(* CODESYS project winhmi.library
   DefaultNamespace: KOSTAL.AF2024.HMI.WinHMI
   DocFormat: reStructuredText
   Description: Interface to WinHMI application
   Author: Martin Hundt
   Title: KOSTAL.AF2024.HMI.WinHMI
   Version: 2.0.0.0
   Company: KOSTAL GmbH & Co.KG
   Placeholder: KOSTAL.AF2024.HMI.WinHMI

Project tree, tasks and I/O mapping:
  libraries: KOSTAL.AF2024.Core.functionResponse, 1.0.0.0 (KOSTAL GmbH & Co.KG); KOSTAL.AF2024.Core.GetSystemTime, 1.0.1.0 (KOSTAL GmbH & Co.KG); KOSTAL.AF2024.Core.ID, 1.0.0.0 (KOSTAL GmbH & Co.KG); KOSTAL.AF2024.Core.JsonTools, 1.0.0.0 (KOSTAL GmbH & Co.KG); KOSTAL.AF2024.Core.ListOf, 1.0.0.0 (KOSTAL GmbH & Co.KG); KOSTAL.AF2024.Core.MainControl, 1.0.0.0 (KOSTAL GmbH & Co.KG); KOSTAL.AF2024.Core.Process, 1.0.999.1 (KOSTAL GmbH & Co.KG); KOSTAL.AF2024.Core.Settings, 1.0.0.0 (KOSTAL GmbH & Co.KG); KOSTAL.AF2024.Core.Station, 1.0.0.0 (KOSTAL GmbH & Co.KG); KOSTAL.AF2024.Core.StringTools, 1.0.0.0 (KOSTAL GmbH & Co.KG); KOSTAL.AF2024.Core.System, 1.0.0.0 (KOSTAL GmbH & Co.KG); KOSTAL.AF2024.Core.Text, 1.0.0.0 (KOSTAL GmbH & Co.KG); KOSTAL.AF2024.HMI.Controls, 1.0.1.0 (KOSTAL GmbH & Co.KG); KOSTAL.AF2024.HMI.I_Hmi, 1.0.0.0 (KOSTAL GmbH & Co.KG); KOSTAL.AF2024.Misc.Counter, 1.0.1.0 (KOSTAL GmbH & Co.KG); Tc2_Standard, 3.4.5.0 (Beckhoff Automation GmbH); Tc2_Utilities, 3.8.2.0 (Beckhoff Automation GmbH); Tc3_JsonXml, 3.4.4.0 (Beckhoff Automation GmbH)
  Aliases/
    data type T_ARTICLESJSON
    data type T_BUTTON_LISTING
    data type T_ExpertPageUserIndex
    data type T_MEDIA_PATH
    data type T_PARAMETERJSON
    data type T_PARAMETERVALUE
  Article/
    data type _ST_Article_FromDevice
    data type _ST_Article_ToDevice
    function block FB_ArticleList [ST]: ActualArticle, AddArticle, Clear, FB_init, FBmain, SelectedArticleName, Set
    interface I_Article: ActualArticle, SelectedArticleName
  Counter/
    data type _ST_Counter_FromDevice
    data type _ST_Counter_ToDevice
    function block FB_Counter [ST]: _HMI_define, ResetEnable
  Listing/
    data type _ST_Listing_FromDevice
    data type _ST_Listing_ToDevice
    function block FB_Page_Listing [ST]: _buttonHandler, _buttonHandler_listing, _listingHandler, _setButton, FB_init, FBmain
  MainControl/
    DUT/
      ListOfIcondition/
        interface I_ListOfCondition: NumberOfMember
        interface I_ListOfCondition_Owner
      data type _E_MainControlMode
      data type _E_MainControlState
    data type _ST_MainControl_FromDevice
    data type _ST_MainControl_toDevice
    function block FB_MainControl [ST]: _buttonHandler, _mainControlHandler, _modeToEnum, _plcStateToEnum, clear, FBmain, ManualDeviceControl
    interface I_MainControl: clear
  Media/
    data type _ST_Media_ToDevice
    function block FB_Media [ST]: Clear, FBmain, SetMedia, ShowMedia, StandardPath
    interface I_Media: Clear, SetMedia, ShowMedia, StandardPath
  Parameters/
    function block _FB_jsonHandler [ST]: Clear, GetJsonString, getValue, ID, NumberOfValues, setValue, Timestamp, _Step_ClearContent, _Step_CreateContent, _Step_ParseContent
    data type _ST_Parameters_FromDevice
    data type _ST_Parameters_ToDevice
    data type E_DataMode
    function block FB_Parameters_Base [ST]: _getParameterValue, _setParameterValue, FullQualifiedFile, ReloadDataFile, _Idle, _readFile, _setParaValue, _HMIdefine, _parameterControl, _resetCondition, FBmain, link_I_getTime
  Project Information/
    function F_GetCompany [ST]
    function F_GetTitle [ST]
    function F_GetVersion [ST]
  Station/
    data type _ST_StationPage_FromDevice
    data type _ST_StationPage_ToDevice
    function block FB_Page_Station [ST]: _buttonHandler, _setButton, _stationHandler, FB_init, FBmain
  Version/
    global variables Global_Version
  XYZ/
    data type _ST_XYZ_FromDevice
    data type _ST_XYZ_ToDevice
    function block FB_page_XYZ [ST]: _buttonHandler, _fillTextLines, _pageHandler, _setButton, FB_init, FBmain
  global variables GVL_CONSTANT
*)

// Aliases/T_ARTICLESJSON
TYPE T_ARTICLESJSON : STRING(6000)
; END_TYPE

// Aliases/T_BUTTON_LISTING
TYPE T_BUTTON_LISTING : WSTRING(3); END_TYPE

// Aliases/T_ExpertPageUserIndex
(*
Description
===========
| Limited data type for the index of an expert page user
*)
TYPE T_ExpertPageUserIndex : INT(0..GVL_CONSTANT.MAX_EXPERT_STATIONS); END_TYPE

// Aliases/T_MEDIA_PATH
TYPE T_MEDIA_PATH : STRING(80)
; END_TYPE

// Aliases/T_PARAMETERJSON
TYPE T_PARAMETERJSON : STRING(6000)
; END_TYPE

// Aliases/T_PARAMETERVALUE
TYPE T_PARAMETERVALUE : STRING(40)
; END_TYPE

// Article/_ST_Article_FromDevice
(*
Description
===========
| Data type to receive article data from WinHMI display
*)
{attribute 'pack_mode' := '1'}
TYPE _ST_Article_FromDevice :
	STRUCT
		SelectedArticleName 	: T_ARTICLENAME;
	END_STRUCT
END_TYPE

// Article/_ST_Article_ToDevice
(*
Description
===========
| Data type to provide article data to WinHMI display
*)
{attribute 'pack_mode' := '1'}
TYPE _ST_Article_ToDevice :
	STRUCT
		ArticleList		: T_ARTICLESJSON;
		ActualArticle 	: T_ARTICLENAME;		(*Shows the actual used Article name	 *)
	END_STRUCT
END_TYPE

// Counter/_ST_Counter_FromDevice
(*
Description
===========
| Data type to provide counter data to WinHMI display
*)
{attribute 'pack_mode' := '1'}
TYPE _ST_Counter_FromDevice :
	STRUCT
		Reset	: BOOL;
	END_STRUCT
END_TYPE

// Counter/_ST_Counter_ToDevice
(*
Description
===========
| Data type to provide counter data to WinHMI display
*)
{attribute 'pack_mode' := '1'}
TYPE _ST_Counter_ToDevice :
	STRUCT
		Passparts		: UDINT;
		Failparts		: UDINT;
		CounterReady 	: BOOL;
		ResetEnable		: BOOL;
	END_STRUCT
END_TYPE

// Listing/_ST_Listing_FromDevice
(*
Description
===========
| Data type to receive listing page data from WinHMI display
*)
{attribute 'pack_mode' := '1'}
TYPE _ST_Listing_FromDevice :
	STRUCT
		IsActive 		: BOOL;		(* 	BOOL	-	Response the state of the Listing Form	 *)
		Button_Left	 	: ARRAY [1..GVL_CONSTANT.LISTING_MAX_LINE] OF BOOL;		(* 	ARRAY[1..10] OF BOOL	-	Status of Button - TRUE = pressed	 *)
		Button_Right	: ARRAY [1..GVL_CONSTANT.LISTING_MAX_LINE] OF BOOL;		(* 	ARRAY[1..10] OF BOOL	-	Status of Button - TRUE = pressed	 *)
	END_STRUCT
END_TYPE

// Listing/_ST_Listing_ToDevice
(*
Description
===========
| Data type to provide listing page data to WinHMI display
*)
{attribute 'pack_mode' := '1'}
TYPE _ST_Listing_ToDevice :
	STRUCT
		
		Activate 		: BOOL;		(* 	BOOL	-	Activate the Listing Form	 *)
		
		Buttons_Left_Active : WORD;		(* 	If bit is TRUE than the correspond Button is visible	 *)
		Buttons_Right_Active : WORD;		(* 	If bit is TRUE than the correspond Button is visible	 *)
		
		Buttons_Left_Text	: ARRAY [1..GVL_CONSTANT.LISTING_MAX_LINE] OF T_BUTTON_LISTING;
		Buttons_Right_Text	: ARRAY [1..GVL_CONSTANT.LISTING_MAX_LINE] OF T_BUTTON_LISTING;
		
		Text 				: ARRAY [1..GVL_CONSTANT.LISTING_MAX_LINE] OF KOSTAL_AF2024_HMI_I_Hmi.T_PAGE_TEXT;	(* Contains the Texts for Line 1..10	 *)
		Status 				: ARRAY [1..GVL_CONSTANT.LISTING_MAX_LINE] OF KOSTAL_AF2024_HMI_I_Hmi.E_STATE;		(* 	Contains the States for Line 1..10	 *)
	END_STRUCT
END_TYPE

// MainControl/DUT/_E_MainControlMode
{attribute 'qualified_only'}
{attribute 'strict'}
TYPE _E_MainControlMode :
(
	undefined := 0,	
	manual,			
	automatic
)USINT;
END_TYPE

// MainControl/DUT/_E_MainControlState
{attribute 'qualified_only'}
{attribute 'strict'}
TYPE _E_MainControlState :
(
	off := 0,	//Power off
	on,			//Power on
	calibrate,	//Power off
	ready,		//Ready to start
	busy,		//running
	finish		//Run empty
)USINT;
END_TYPE

// MainControl/_ST_MainControl_FromDevice
(*
Description
===========
| Data type to receive Main Control data from WinHMI display
*)
{attribute 'pack_mode' := '1'}
TYPE _ST_MainControl_FromDevice :
	STRUCT
		Language 			: T_LANGUAGENAME;		(* 	STRING(40)	- Selected Languagename	 *)
				
		Button_Auto 		: BOOL;		(* 	BOOL	- Status of Button - TRUE = pressed	 *)
		Button_Manual : BOOL;		(* 	BOOL	- Status of Button - TRUE = pressed	 *)
		Button_Door 		: BOOL;		(* 	BOOL	- Status of Button - TRUE = pressed	 *)

		Button_OnOff 		: BOOL;		(* BOOL *)
		Button_StartStop : BOOL;		(* BOOL *)
		Button_workEmpty : BOOL;		(* BOOL *)
		
		UserLevel	: BYTE; 	//operator = 0, service = 1, quality = 2

	END_STRUCT
END_TYPE

// MainControl/_ST_MainControl_toDevice
(*
Description
===========
| Data type to provide Main Control data to WinHMI display
*)
{attribute 'pack_mode' := '1'}
TYPE _ST_MainControl_toDevice :
	STRUCT
		Status_Auto 	: BOOL;		(* 	BOOL	-	If TRUE > Text "Auto" has a yellow background	 *)
		Status_Manual : BOOL;		(* 	BOOL	-	If TRUE > Text "Manual" has a yellow background	 *)
	
		Status_Door_Close : BOOL;		(* 	BOOL	-	If TRUE > Text "Door" has a blue background	 *)
		Status_Door_Open 	: BOOL;		(* 	BOOL	-	If TRUE > Text "Door" has a red background	 *)
		Status_Door_Safe 	: BOOL;		(* 	BOOL	-	If TRUE > Text "Door" has a green background	 *)

		Manual_Enable 	: BOOL;		(* 	BOOL	-	If TRUE > Button in bottom of Text "Manual" is visible	 *)
		Parameters_Enable 		: BOOL;		(* 	BOOL	-	If TRUE > Button in bottom of Text "Data" is visible	 *)
		Auto_Enable 		: BOOL;		(* 	BOOL	-	If TRUE > Button in bottom of Text "Auto" is visible	 *)
		Door_Enable 		: BOOL;		(* 	BOOL	-	If TRUE > Button in bottom of Text "Door" is visible	 *)
		Article_Enable 	: BOOL;		(* 	BOOL	-	If TRUE > Button in bottom of Text "Article" is visible	 *)

		(*  Buttons *)
		OnOff_Enable	: BOOL;
		RunStop_Enable	: BOOL;
		RunEmpty_Enable 	: BOOL;
		
		Status_On 		: BOOL;		(* BOOL *)
		Status_Run 		: BOOL;		(* BOOL *)
		Status_RunEmpty 	: BOOL;		(* BOOL *)
		ManualDeviceControl_Enable	: BOOL;
		
		//main Control
		State		: USINT;
		Mode		: USINT;
				
	END_STRUCT
END_TYPE

// Media/_ST_Media_ToDevice
(*
Description
===========
| Data type to provide article data to WinHMI display
*)
{attribute 'pack_mode' := '1'}
TYPE _ST_Media_ToDevice :
	STRUCT
		MediaAddress		: T_MEDIA_PATH;
	END_STRUCT
END_TYPE

// Parameters/_ST_Parameters_FromDevice
(*
Description
===========
| Data type to receive parameter data from WinHMI display
*)
{attribute 'pack_mode' := '1'}
TYPE _ST_Parameters_FromDevice :
	STRUCT
		SelectedParameter 			: BYTE;		(* 	BYTE	- Selected Dataset 	 *)
		NewValue 				: T_PARAMETERVALUE;		(* 	STRING(40)	-	New Data value	 *)
		NewValueTransmit 	: BOOL;		(* 	BOOL	-	New value is valid	 *)

	END_STRUCT
END_TYPE

// Parameters/_ST_Parameters_ToDevice
(*
Description
===========
| Data type to provide XYZ page parameter data to WinHMI display
*)
{attribute 'pack_mode' := '1'}
TYPE _ST_Parameters_ToDevice :
	STRUCT
		ParameterValuesJson		: T_PARAMETERJSON;
		NewValueAccept			: BOOL;
	END_STRUCT
END_TYPE

// Parameters/E_DataMode
{attribute 'qualified_only'}
{attribute 'strict'}
TYPE E_DataMode :
(
	Idle := 0,
	ReadFile,
	WriteParameter
);
END_TYPE

// Station/_ST_StationPage_FromDevice
(*
Description
===========
| Data type to receive 3D page from WinHMI display
*)
{attribute 'pack_mode' := '1'}
TYPE _ST_StationPage_FromDevice :
	STRUCT
		Button_F1 : BOOL;		(* 	BOOL	- Status of Button - TRUE = pressed	 *)
		Button_F2 : BOOL;		(* 	BOOL	- Status of Button - TRUE = pressed	 *)
		Button_F3 : BOOL;		(* 	BOOL	- Status of Button - TRUE = pressed	 *)
		Button_F4 : BOOL;		(* 	BOOL	- Status of Button - TRUE = pressed	 *)
		Button_F5 : BOOL;		(* 	BOOL	- Status of Button - TRUE = pressed	 *)
		Button_F6 : BOOL;		(* 	BOOL	- Status of Button - TRUE = pressed	 *)
		Button_F7 : BOOL;		(* 	BOOL	- Status of Button - TRUE = pressed	 *)

		Button_On 			: BOOL;		(* 	BOOL	- Status of Button - TRUE = pressed	 *)
		Button_Minus 	: BOOL;		(* 	BOOL	- Status of Button - TRUE = pressed	 *)
		Button_Enter 	: BOOL;		(* 	BOOL	- Status of Button - TRUE = pressed	 *)
		Button_Plus 		: BOOL;		(* 	BOOL	- Status of Button - TRUE = pressed	 *)
		Button_Escape 	: BOOL;		(* 	BOOL	- Status of Button - TRUE = pressed	 *)

	END_STRUCT
END_TYPE

// Station/_ST_StationPage_ToDevice
(*
Description
===========
| Data type to provide station page data to WinHMI display
*)
{attribute 'pack_mode' := '1'}
TYPE _ST_StationPage_ToDevice :
	STRUCT

		StationName : KOSTAL_AF2024_HMI_I_Hmi.T_PAGE_TEXT;			(* Response the requested Username during Initialization	 *)
		
		TextLines : ARRAY [1..3] OF KOSTAL_AF2024_HMI_I_Hmi.T_PAGE_TEXT;		(* 	Four Textlines  *)

		HmiState	: KOSTAL_AF2024_HMI_I_HMI.E_STATE;

		F1_Text 	: KOSTAL_AF2024_HMI_I_HMI.T_F_BUTTON_TEXT ;		(* 	If not empty the Button is visible with Text *)
		F2_Text 	: KOSTAL_AF2024_HMI_I_HMI.T_F_BUTTON_TEXT ;		(* 	If not empty the Button is visible with Text *)
		F3_Text 	: KOSTAL_AF2024_HMI_I_HMI.T_F_BUTTON_TEXT ;		(* 	If not empty the Button is visible with Text *)
		F4_Text 	: KOSTAL_AF2024_HMI_I_HMI.T_F_BUTTON_TEXT ;		(* 	If not empty the Button is visible with Text *)
		F5_Text 	: KOSTAL_AF2024_HMI_I_HMI.T_F_BUTTON_TEXT ;		(* 	If not empty the Button is visible with Text *)
		F6_Text 	: KOSTAL_AF2024_HMI_I_HMI.T_F_BUTTON_TEXT ;		(* 	If not empty the Button is visible with Text *)
		F7_Text 	: KOSTAL_AF2024_HMI_I_HMI.T_F_BUTTON_TEXT ;		(* 	If not empty the Button is visible with Text *)
                                                                                                                    
		On_Text 	: KOSTAL_AF2024_HMI_I_HMI.T_BUTTON_TEXT;		(* 	If not empty the Button is visible with Text *)
		Minus_Text 	: KOSTAL_AF2024_HMI_I_HMI.T_BUTTON_TEXT;		(* 	If not empty the Button is visible with Text *)
		Enter_Text 	: KOSTAL_AF2024_HMI_I_HMI.T_BUTTON_TEXT;		(* 	If not empty the Button is visible with Text *)
		Plus_Text 	: KOSTAL_AF2024_HMI_I_HMI.T_BUTTON_TEXT;		(* 	If not empty the Button is visible with Text *)
		Escape_Text : KOSTAL_AF2024_HMI_I_HMI.T_BUTTON_TEXT;		(* 	If not empty the Button is visible with Text *)

		//IsValidUser	: BOOL; (* TRUE if a valid user is linked *)
	END_STRUCT
END_TYPE

// XYZ/_ST_XYZ_FromDevice
(*
Description
===========
| Data type to receive XYZ page data from WinHMI display
*)
{attribute 'pack_mode' := '1'}
TYPE _ST_XYZ_FromDevice :
	STRUCT
		
		Button_Forward 	: BOOL;		(* 	BOOL	- Status of Button - TRUE = pressed	 *)
		Button_Backward	: BOOL;		(* 	BOOL	- Status of Button - TRUE = pressed	 *)
		Button_Right 	: BOOL;		(* 	BOOL	- Status of Button - TRUE = pressed	 *)
		Button_Left 		: BOOL;		(* 	BOOL	- Status of Button - TRUE = pressed	 *)
		Button_Up 		: BOOL;		(* 	BOOL	- Status of Button - TRUE = pressed	 *)
		Button_Down 		: BOOL;		(* 	BOOL	- Status of Button - TRUE = pressed	 *)		
		Button_Custom_1 		: BOOL;		(* 	BOOL	- Status of Button - TRUE = pressed	 *)
		Button_Custom_2 	: BOOL;		(* 	BOOL	- Status of Button - TRUE = pressed	 *)
		Button_Custom_3 	: BOOL;		(* 	BOOL	- Status of Button - TRUE = pressed	 *)
		Button_Custom_4 	: BOOL;		(* 	BOOL	- Status of Button - TRUE = pressed	 *)
		Button_StepPlus 	: BOOL;		(* 	BOOL	- Status of Button - TRUE = pressed	 *)
		Button_StepMinus : BOOL;		(* 	BOOL	- Status of Button - TRUE = pressed	 *)
		Button_Off 		: BOOL;		(* 	BOOL	- Status of Button - TRUE = pressed	 *)

	END_STRUCT
END_TYPE

// XYZ/_ST_XYZ_ToDevice
(*
Description
===========
| Data type to provide XYZ page data to WinHMI display
*)
{attribute 'pack_mode' := '1'}
TYPE _ST_XYZ_ToDevice :
	STRUCT
		Activate 			: BOOL;		(* 	BOOL	-	If TRUE > Form to handle 3Dimension Function (Axis)	 *)

		Text 			: ARRAY [1..4] OF T_PAGE_TEXT;		(* Four Textlines from 3Dimension Form	 *)
		
		Button_Custom1_Text 		: KOSTAL_AF2024_HMI_I_Hmi.T_F_BUTTON_TEXT;		(* If nor empty the Button is visible with Text*)
		Button_Custom2_Text 		: KOSTAL_AF2024_HMI_I_Hmi.T_F_BUTTON_TEXT;		(* If nor empty the Button is visible with Text*)
		Button_Custom3_Text 		: KOSTAL_AF2024_HMI_I_Hmi.T_F_BUTTON_TEXT;		(* If nor empty the Button is visible with Text*)
		Button_Custom4_Text 		: KOSTAL_AF2024_HMI_I_Hmi.T_F_BUTTON_TEXT;		(* If nor empty the Button is visible with Text*)
		
		Button_Forward_Active 	: BOOL;		 
		Button_Backward_Active	: BOOL;		 
		Button_Right_Active 		: bool;		 
		Button_Left_Active 		: BOOL;	
		Button_Up_Active 		: BOOL;		 
		Button_Down_Active		: bool;	
	 	Button_Plus_Text 		: KOSTAL_AF2024_HMI_I_Hmi.T_F_BUTTON_TEXT;		(* 	STRING(10)	-	If nor empty the Button is visible with Text in upper position	 *)
		Button_Minus_Text 		: KOSTAL_AF2024_HMI_I_Hmi.T_F_BUTTON_TEXT;		(* 	STRING(10)	-	If nor empty the Button is visible with Text in upper position	 *)	
END_STRUCT
END_TYPE

// Version/Global_Version
{attribute 'TcGenerated'}
{attribute 'no-analysis'}
{attribute 'linkalways'}
// This function has been automatically generated from the project information.
VAR_GLOBAL CONSTANT
	{attribute 'const_non_replaced'}
	stLibVersion_KOSTAL_AF2024_HMI_WinHMI : ST_LibVersion := (iMajor := 2, iMinor := 0, iBuild := 0, iRevision := 0, nFlags := 0, sVersion := '2.0.0.0');
END_VAR

// GVL_CONSTANT
{attribute 'qualified_only'}
VAR_GLOBAL CONSTANT

	PAGE_STATION_TEXT_MAX_LINE	: INT:= 4;	//INT:= 4	Maximum number of main page lines
	
	LISTING_MAX_LINE		: INT:= 10;	//INT:= 10	Maximum number of lines on listing page

	EXPERTUSERS_MAX_NUMBER	: UINT:= 32;	// UINT:= 26 - define max user number from Array[1..26]
	MAX_EXPERT_STATIONS 		: INT := 32;
	
	MAX_ARTICLES			: UINT := 120;
END_VAR

// Article/FB_ArticleList
(*

:Author: Martin Hundt <m.hundt@kostal.com>
:Date: 2021-08-16

Function
========
*)
FUNCTION_BLOCK PUBLIC FB_ArticleList IMPLEMENTS I_Article


VAR

	//****************************************************************************
	//Connector
	//****************************************************************************
	{attribute 'Article_2024_V0'}
	_connector_FROM_Device	: _ST_Article_FromDevice;	//ST_ARTICLE_FROMDEVICE
	_connector_TO_Device	: _ST_Article_ToDevice;		//ST_ARTICLE_TODEVICE
	//****************************************************************************
	//****************************************************************************

	//_articleList				: FB_ArticleList;
	
	_articleList	: KOSTAL_AF2024_Core_ListOf.FB_ListOfString_UTF8;
	_json	: T_PARAMETERJSON;
	_isSet	: BOOL;	//Avoid setting the same list again to reduce system load

	
END_VAR

(*
Description
===========
| Name of currently selected article
*)
PROPERTY PUBLIC ActualArticle : T_ARTICLENAME
SET

_connector_TO_Device.ActualArticle := ActualArticle;
END_SET
END_PROPERTY

(*
Description
===========
| Add article to article list
*)
METHOD PUBLIC AddArticle : BOOL;
VAR_INPUT
	Name		: KOSTAL_AF2024_Core_Settings.T_MaxString_UTF8;
	Response	: KOSTAL_AF2024_Core_functionResponse.I_T_functionResponse_Owner;
END_VAR

VAR
	_response	: KOSTAL_AF2024_Core_functionResponse.T_functionResponse;
END_VAR
IF Name = '' THEN 
	_response.success := FALSE;
	_response.status := "Article name is empty";
ELSIF NOT _articleList.addLine(Name) THEN
	_response.success := FALSE;
	_response.status := "Article list is full";
ELSE
	AddArticle := TRUE;
	_response.success := TRUE;
	_isSet := FALSE;
END_IF

IF Response <> 0 THEN
	Response.success := _response.success;
	Response.status := _response.status;
END_IF
END_METHOD

(*
Description
===========
| Clear article list
*)
METHOD Clear
VAR_INPUT
END_VAR
_articleList.clear();
_isSet := false;
END_METHOD

METHOD FB_init : BOOL
VAR_INPUT
	bInitRetains : BOOL; // if TRUE, the retain variables are initialized (warm start / cold start)
	bInCopyCode : BOOL;  // if TRUE, the instance afterwards gets moved into the copy code (online change)
END_VAR
//Set maximum number of articles according to maximum JSON string lenght

_articleList.maxLine := (SIZEOF(T_PARAMETERJSON) - 14)/16;
END_METHOD

METHOD PUBLIC FBmain : BOOL
_connector_TO_Device.ArticleList := _json;
END_METHOD

(*
Description
===========
| Name of currently selected article
*)
PROPERTY PUBLIC SelectedArticleName : T_ARTICLENAME
GET
 SelectedArticleName := _connector_FROM_Device.SelectedArticleName;
END_GET
END_PROPERTY

(*
Description
===========
| Set the created article List to HMI
*)
METHOD Set

//VAR_INPUT
//	Response	: KOSTAL_AF2024_Core_functionResponse.I_T_functionResponse_Owner;
//END_VAR


VAR
	_parser : Tc3_JsonXml.FB_JsonDomParser;
	jsonDoc		: SJsonValue;
	jsonArray	: SJsonValue;
	_i	: UDINT;
	_value	: STRING;
	
	_response	: KOSTAL_AF2024_Core_functionResponse.I_T_functionResponse_Owner;
END_VAR
IF _isSet THEN RETURN; END_IF


jsonDoc := _parser.NewDocument();

jsonArray := _parser.AddArrayMember(jsonDoc, 'CONTENT',0);

FOR _i:=1 TO _articleList.NumberOfLines DO
	_value := _articleList.line_GET(_i);
	_parser.PushbackStringValue(jsonArray, _value);
END_FOR



_parser.CopyDocument(_json, SIZEOF(T_ARTICLESJSON));

_isSet := TRUE;
END_METHOD

END_FUNCTION_BLOCK

// Article/I_Article
(*
Description
===========
| Application interface for article page
*)
INTERFACE I_Article

(*
Description
===========
| Name of currently selected article
*)
PROPERTY PUBLIC ActualArticle : T_ARTICLENAME
SET
END_SET
END_PROPERTY

(*
Description
===========
| Name of currently selected article
*)
PROPERTY PUBLIC SelectedArticleName : T_ARTICLENAME
GET
END_GET
END_PROPERTY

END_INTERFACE

// Counter/FB_Counter
FUNCTION_BLOCK FB_Counter EXTENDS KOSTAL_AF2024_Misc_Counter._FB_Base

VAR

	

	
	//===========================================================================================================
	//Interfaces
	//===========================================================================================================

	
	//****************************************************************************
	//Connector
	//****************************************************************************
		{attribute 'Counter_2024_V0'}
	_connector_TO_Device	: _ST_Counter_ToDevice;
	_connector_FROM_Device	: _ST_Counter_FromDevice;	
	//****************************************************************************
	
	_Hmi_station		: FB_Page_Station;
	
	

END_VAR

METHOD PROTECTED _HMI_define
VAR_INPUT
END_VAR

_pageStation := _Hmi_station;
_Hmi_station.FBmain();

SUPER^._HMI_define();

//Counter
IF _Istorage = 0 THEN
	_connector_TO_Device.Failparts := _connector_TO_Device.Failparts := 0;
	RETURN;
END_IF

IF _connector_FROM_Device.Reset THEN
	_counterFail.Init(0);
	_counterPass.Init(0);
END_IF
_connector_TO_Device.Failparts := _counterFail.Counter;
_connector_TO_Device.Passparts := _counterPass.Counter;
_connector_TO_Device.CounterReady:= _Istorage.State.ready AND _initFromStorageDone;
_connector_TO_Device.ResetEnable := _resetEnable;
END_METHOD

//Set true to enable reset button on HMI
PROPERTY ResetEnable : BOOL
GET
ResetEnable := _resetEnable;
END_GET
SET
_resetEnable := ResetEnable;
END_SET
END_PROPERTY

END_FUNCTION_BLOCK

// Station/FB_Page_Station
(*

:Author: Martin Hundt <m.hundt@kostal.com>
:Date: 2020-03-09

Function
========
Interface for WinHMI Station Page

Usage
=====
See best practice samples and documentation

*)
FUNCTION_BLOCK PUBLIC FB_Page_Station EXTENDS KOSTAL_AF2024_HMI_I_Hmi.FB_Page_Station


VAR

	//****************************************************************************
	//Connector
	//****************************************************************************
	{attribute 'Page_Station_2024_V0'}
	_connector_FROM_Device		: _ST_StationPage_FromDevice;	
	_connector_TO_Device		: _ST_StationPage_ToDevice;		
	//****************************************************************************
	//****************************************************************************



	
	_pulse_on		: F_TRIG;	
	_pulse_minus	: F_TRIG;	
	_pulse_enter	: F_TRIG;	
	_pulse_plus	: F_TRIG;	
	_pulse_escape	: F_TRIG;	
          
	_pulse_F	: ARRAY[1..7] OF F_TRIG;	

END_VAR

METHOD PROTECTED _buttonHandler : BOOL
VAR_INPUT
END_VAR

VAR
	_index: INT;	// INT
END_VAR
_pulse_on			(CLK:= _connector_FROM_Device.Button_On);
_pulse_minus	(CLK:= _connector_FROM_Device.Button_Minus);
_pulse_enter	(CLK:= _connector_FROM_Device.Button_Enter);
_pulse_plus		(CLK:= _connector_FROM_Device.Button_Plus);
_pulse_escape	(CLK:= _connector_FROM_Device.Button_Escape);
      
_pulse_F[1](CLK:= _connector_FROM_Device.Button_F1);
_pulse_F[2](CLK:= _connector_FROM_Device.Button_F2);
_pulse_F[3](CLK:= _connector_FROM_Device.Button_F3);
_pulse_F[4](CLK:= _connector_FROM_Device.Button_F4);
_pulse_F[5](CLK:= _connector_FROM_Device.Button_F5);
_pulse_F[6](CLK:= _connector_FROM_Device.Button_F6);
_pulse_F[7](CLK:= _connector_FROM_Device.Button_F7);
END_METHOD

METHOD PROTECTED _setButton : WSTRING

VAR_INPUT
	control	: KOSTAL_AF2024_HMI_Controls.I_T_Button_controlled;	//KOSTAL_TC3_Controls_button.FB_Button_controlled
END_VAR

IF control.Visible THEN

	IF control.Text = "" THEN
		_setButton:= " ";
	ELSE
		_setButton:= control.Text;
	END_IF

ELSE

	_setButton:= "";

END_IF
END_METHOD

METHOD PROTECTED _stationHandler
VAR_INPUT
END_VAR

VAR
	_index: INT;	// INT
END_VAR
//TO
//hmiState (replaces status)
IF _status.isError() THEN
	_connector_TO_Device.HmiState := KOSTAL_AF2024_HMI_I_HMI.E_STATE.ERROR;
ELSIF _status.isFail() THEN
	_connector_TO_Device.HmiState := KOSTAL_AF2024_HMI_I_HMI.E_STATE.FAIL;
ELSIF _status.isPass() THEN
	_connector_TO_Device.HmiState := KOSTAL_AF2024_HMI_I_HMI.E_STATE.PASS;
ELSIF _status.isMessage() OR  _status.isMasterMessage() THEN
	_connector_TO_Device.HmiState := KOSTAL_AF2024_HMI_I_HMI.E_STATE.ATTENTION;
//ELSIF _status.isText() THEN
//	_connector_TO_Device.HmiState := KOSTAL_AF2024_HMI_I_HMI.E_STATE.PASS;
ELSE
	_connector_TO_Device.HmiState := KOSTAL_AF2024_HMI_I_HMI.E_STATE.NONE;
END_IF



//
_connector_TO_Device.Enter_Text:= 	_setButton(_Enter);
_connector_TO_Device.Escape_Text:=	_setButton(_Escape);
_connector_TO_Device.On_Text:= 		_setButton(_OnOff);
_connector_TO_Device.Minus_Text:=	_setButton(_Minus);
_connector_TO_Device.Plus_Text:= 	_setButton(_Plus);

//F(1..7)
_connector_TO_Device.F1_Text:= 		_setButton(_custom.Button(1));
_connector_TO_Device.F2_Text:= 		_setButton(_custom.Button(2));
_connector_TO_Device.F3_Text:= 		_setButton(_custom.Button(3));
_connector_TO_Device.F4_Text:= 		_setButton(_custom.Button(4));
_connector_TO_Device.F5_Text:= 		_setButton(_custom.Button(5));
_connector_TO_Device.F6_Text:= 		_setButton(_custom.Button(6));
_connector_TO_Device.F7_Text:= 		_setButton(_custom.Button(7));
//F8 is handled internal by VB

_connector_TO_Device.StationName	:= _name;
_connector_TO_Device.TextLines[1]:= _text.line_01;
_connector_TO_Device.TextLines[2]:= _text.line_02;
_connector_TO_Device.TextLines[3]:= _text.line_03;



//FROM

_onOff.Sign		:= _connector_FROM_Device.Button_On;
_onOff.Pulse	:= _pulse_on.Q;
      
_minus.Sign		:= _connector_FROM_Device.Button_Minus;
_minus.Pulse	:= _pulse_minus.Q;
IF _onOff.Pulse THEN
	_index := _index+1;
END_IF
      
_enter.Sign		:= _connector_FROM_Device.Button_Enter;
_enter.Pulse	:= _pulse_enter.Q;
      
_plus.Sign		:= _connector_FROM_Device.Button_Plus;
_plus.Pulse	:= _pulse_plus.Q;
      
_escape.Sign		:= _connector_FROM_Device.Button_Escape;
_escape.Pulse	:= _pulse_escape.Q;
      
_custom.Button_Owner(1).Sign		:= _connector_FROM_Device.Button_F1;
_custom.Button_Owner(1).Pulse	:= _pulse_F[1].Q;

_custom.Button_Owner(2).Sign		:= _connector_FROM_Device.Button_F2;
_custom.Button_Owner(2).Pulse	:= _pulse_F[2].Q;

_custom.Button_Owner(3).Sign		:= _connector_FROM_Device.Button_F3;
_custom.Button_Owner(3).Pulse	:= _pulse_F[3].Q;

_custom.Button_Owner(4).Sign		:= _connector_FROM_Device.Button_F4;
_custom.Button_Owner(4).Pulse	:= _pulse_F[4].Q;
 
_custom.Button_Owner(5).Sign		:= _connector_FROM_Device.Button_F5;
_custom.Button_Owner(5).Pulse	:= _pulse_F[5].Q;

_custom.Button_Owner(6).Sign		:= _connector_FROM_Device.Button_F6;
_custom.Button_Owner(6).Pulse	:= _pulse_F[6].Q;

_custom.Button_Owner(7).Sign		:= _connector_FROM_Device.Button_F7;
_custom.Button_Owner(7).Pulse	:= _pulse_F[7].Q;
END_METHOD

(*
Description
===========
| Method is called automatically
| Do not call manually
*)
METHOD FB_init : BOOL
VAR_INPUT
	bInitRetains : BOOL; // if TRUE, the retain variables are initialized (warm start / cold start)
	bInCopyCode : BOOL;  // if TRUE, the instance afterwards gets moved into the copy code (online change)
END_VAR

VAR
	_index	: INT;	//INT
	x: BOOL;
END_VAR
END_METHOD

METHOD PUBLIC FBmain : BOOL
VAR_INPUT
END_VAR

VAR
END_VAR
_buttonHandler();
_stationHandler();
END_METHOD

END_FUNCTION_BLOCK

// Listing/FB_Page_Listing
(*

:Author: Martin Hundt <m.hundt@kostal.com>
:Date: 2020-03-09

Function
========
Interface for WinHMI Listing Page

Usage
=====
See best practice samples and documentation

*)
FUNCTION_BLOCK PUBLIC FB_Page_Listing EXTENDS KOSTAL_AF2024_HMI_I_Hmi.FB_Page_Listing


VAR

	//****************************************************************************
	//Connector
	//****************************************************************************
	
	{attribute 'Page_Listing_2024_V0'}
	_connector_FROM_Device	: _ST_Listing_FromDevice;	//ST_LISTING_FROMDEVICE
	_connector_TO_Device	: _ST_Listing_ToDevice;		//ST_LISTING_TODEVICE
	//****************************************************************************
	//****************************************************************************

	
	
	//page Listing

	_pulse_buttons_Left		: ARRAY[1..KOSTAL_AF2024_HMI_I_HMI.GVL_CONSTANT.MAX_LISTING_LINE] OF F_TRIG;	
	_pulse_buttons_Right	: ARRAY[1..KOSTAL_AF2024_HMI_I_HMI.GVL_CONSTANT.MAX_LISTING_LINE] OF F_TRIG;	
	
	
	
END_VAR

METHOD PROTECTED _buttonHandler
VAR_INPUT
END_VAR
_buttonHandler_listing();
END_METHOD

METHOD PROTECTED _buttonHandler_listing : BOOL
VAR_INPUT
END_VAR

VAR
	_index: INT;	// INT
END_VAR

FOR _index:= 1 TO KOSTAL_AF2024_HMI_I_HMI.GVL_CONSTANT.MAX_LISTING_LINE DO
	_pulse_buttons_Left[_index]	(CLK:= _connector_FROM_Device.Button_Left[_index]);
	_pulse_buttons_Right[_index]	(CLK:= _connector_FROM_Device.Button_Right[_index]);
END_FOR
END_METHOD

METHOD PROTECTED _listingHandler
VAR_INPUT
END_VAR

VAR
	_index: INT;	// INT
	
END_VAR
//TO
_connector_TO_Device.Activate := _activate AND NOT _deactivate;

_connector_TO_Device.Buttons_Left_Active := 0;
_connector_TO_Device.Buttons_Right_Active := 0;
	

FOR _index:= 1 TO KOSTAL_AF2024_HMI_I_HMI.GVL_CONSTANT.MAX_LISTING_LINE DO
	
	_connector_TO_Device.Text[_index]		:= THIS^._messages.Message(_index).Content;
	_connector_TO_Device.Status[_index]		:= 	THIS^._messages.Message(_index).State;
	
	_connector_TO_Device.Buttons_Left_Active := _connector_TO_Device.Buttons_Left_Active + SHL(BOOL_TO_WORD(THIS^._Buttons.Button_Left(_index).Visible), _index - 1);
	_connector_TO_Device.Buttons_Right_Active := _connector_TO_Device.Buttons_Right_Active + SHL(BOOL_TO_WORD(THIS^._Buttons.Button_Right(_index).Visible), _index - 1);
	
	_connector_TO_Device.Buttons_Left_Text[_index] := _Buttons.Button_Left(_index).Text;
	_connector_TO_Device.Buttons_Right_Text[_index] := _Buttons.Button_Right(_index).Text;


END_FOR


//FROM

FOR _index:= 1 TO KOSTAL_AF2024_HMI_I_HMI.GVL_CONSTANT.MAX_LISTING_LINE DO

	THIS^._Buttons.Button_Left_Owner(_index).Sign	:= _connector_FROM_Device.Button_Left[_index];
	THIS^._Buttons.Button_Left_Owner(_index).Pulse	:= _pulse_buttons_Left[_index].Q;
           
	THIS^._Buttons.Button_Right_Owner(_index).Sign	:= _connector_FROM_Device.Button_Right[_index];
	THIS^._Buttons.Button_Right_Owner(_index).Pulse	:= _pulse_buttons_Right[_index].Q;

END_FOR

_isActiv	:= _connector_FROM_Device.IsActive;
END_METHOD

METHOD PROTECTED _setButton : WSTRING

VAR_INPUT
	control	: KOSTAL_AF2024_HMI_Controls.T_Button_controlled;	//KOSTAL_TC3_Controls_button.FB_Button_controlled
END_VAR

IF control.Visible THEN

	IF control.Text = "" THEN
		_setButton:= " ";
	ELSE
		_setButton:= control.Text;
	END_IF

ELSE

	_setButton:= "";

END_IF
END_METHOD

(*
Description
===========
| Method is called automatically
| Do not call manually
*)
METHOD FB_init : BOOL
VAR_INPUT
	bInitRetains : BOOL; // if TRUE, the retain variables are initialized (warm start / cold start)
	bInCopyCode : BOOL;  // if TRUE, the instance afterwards gets moved into the copy code (online change)
END_VAR

VAR
	_index	: INT;	//INT
	x: BOOL;
END_VAR
END_METHOD

METHOD PUBLIC FBmain : BOOL
VAR_INPUT
END_VAR

VAR
END_VAR
_buttonHandler();

_listingHandler();
END_METHOD

END_FUNCTION_BLOCK

// MainControl/DUT/ListOfIcondition/I_ListOfCondition
(*
	Read-Only access to List
*)
INTERFACE I_ListOfCondition EXTENDS KOSTAL_AF2024_Core_ListOf._I_Interface_Base

(*
	Return the number of members in List
*)
PROPERTY PUBLIC NumberOfMember : UDINT
GET
END_GET
END_PROPERTY

END_INTERFACE

// MainControl/DUT/ListOfIcondition/I_ListOfCondition_Owner
(*
	full access to List
*)
INTERFACE I_ListOfCondition_Owner EXTENDS KOSTAL_AF2024_Core_ListOf._I_Interface_Base_Owner

END_INTERFACE

// MainControl/FB_MainControl
(*

:Author: Martin Hundt <m.hundt@kostal.com>
:Date: 2020-03-09

Function
========
WinHMI MainControl interface

Usage
=====
See best practice samples and documentation

*)
FUNCTION_BLOCK PUBLIC FB_MainControl EXTENDS KOSTAL_AF2024_HMI_I_Hmi.FB_MainControl IMPLEMENTS I_MainControl


VAR

	//****************************************************************************
	//Connector
	//****************************************************************************
	{attribute 'MainControl_2024_V0'}
	_connector_FROM_Device	: _ST_MainControl_FROMDEVICE;	
	_connector_TO_Device	: _ST_MainControl_toDevice;		
	//****************************************************************************
	//****************************************************************************

	_manualDeviceControl	: BOOL;

	_pulse_onOff		: F_TRIG;	
	_pulse_startStop	: F_TRIG;	
	_pulse_workEmpty	: F_TRIG;	        
	_pulse_manual		: F_TRIG;	
	_pulse_auto			: F_TRIG;
	_pulse_door			: F_TRIG;	
	
	
	
END_VAR

VAR CONSTANT
	
END_VAR

METHOD PROTECTED _buttonHandler : BOOL
VAR_INPUT
END_VAR

VAR
	_index: INT;	// INT
END_VAR
_pulse_onOff			(CLK:= _connector_FROM_Device.Button_OnOff);
_pulse_startStop	(CLK:= _connector_FROM_Device.Button_StartStop);
_pulse_workEmpty	(CLK:= _connector_FROM_Device.Button_workEmpty);
       
_pulse_manual	(CLK:= _connector_FROM_Device.Button_Manual);
_pulse_auto		(CLK:= _connector_FROM_Device.Button_Auto);
_pulse_door		(CLK:= _connector_FROM_Device.Button_Door);
END_METHOD

METHOD PROTECTED _mainControlHandler : BOOL

VAR

	_index: INT;	// INT
	
END_VAR

//TO
_connector_TO_Device.Auto_Enable	:= _Auto.Visible;
_connector_TO_Device.Parameters_Enable	:= _Parameters.Visible;

_connector_TO_Device.Manual_Enable	:= _Manual.Visible;

_connector_TO_Device.Door_Enable				:=	_Door.Visible;
_connector_TO_Device.Status_Door_Close	:= 	_statusDoor_close AND NOT _statusDoor_safe;
_connector_TO_Device.Status_Door_Open		:= 	_statusDoor_open;
_connector_TO_Device.Status_Door_Safe	:= 	_statusDoor_safe;

_connector_TO_Device.Article_Enable	:= _Article.Visible;


_connector_TO_Device.OnOff_Enable		:= 	_OnOff.Visible;
_connector_TO_Device.RunStop_Enable		:= 	_runStop.Visible;
_connector_TO_Device.RunEmpty_Enable	:=	_RunEmpty.Visible;

_connector_TO_Device.ManualDeviceControl_Enable := _manualDeviceControl AND _mainControl.Mode.manual;

//State and mode
_connector_TO_Device.State 		:= _plcStateToEnum(_mainControl.Demand);
_connector_TO_Device.Status_On			:= 	NOT _mainControl.Demand.PowerOff;
_connector_TO_Device.Status_Run			:= 	_mainControl.Demand.Run OR _mainControl.Demand.RunToHome;
_connector_TO_Device.Status_RunEmpty		:= 	_mainControl.RunEmpty;

_connector_TO_Device.Mode			:= _modeToEnum(_mainControl.Mode);
_connector_TO_Device.Status_Manual		:= _mainControl.Mode.manual;
_connector_TO_Device.Status_Auto		:= _mainControl.Mode.automatic;

//FROM

_Auto.Sign		:=	_connector_FROM_Device.Button_Auto;
_Auto.Pulse	:= _pulse_auto.Q;

_Manual.Sign		:=	_connector_FROM_Device.Button_Manual;
_Manual.Pulse	:= _pulse_manual.Q;


_Door.Sign		:=	_connector_FROM_Device.Button_Door;
_Door.Pulse	:= _pulse_door.Q;

_OnOff.Sign		:=	_connector_FROM_Device.Button_OnOff;
_OnOff.Pulse	:= _pulse_onOff.Q;

_RunStop.Sign		:=	_connector_FROM_Device.Button_StartStop;
_RunStop.Pulse	:= _pulse_startStop.Q;

_RunEmpty.Sign		:=	_connector_FROM_Device.Button_workEmpty;
_RunEmpty.Pulse	:= _pulse_workEmpty.Q;
     
_Language			:= _connector_FROM_Device.Language;


CASE _connector_FROM_Device.UserLevel OF
	1:	_UserLevel := KOSTAL_AF2024_HMI_I_HMI.E_UserLevel.service;
	2:	_UserLevel := KOSTAL_AF2024_HMI_I_HMI.E_UserLevel.quality;
ELSE
	_UserLevel := KOSTAL_AF2024_HMI_I_HMI.E_UserLevel.operator;
END_CASE
END_METHOD

METHOD PROTECTED _modeToEnum : _E_MainControlMode
VAR_INPUT
	mode	: KOSTAL_AF2024_Core_process.I_T_processMode;
END_VAR
IF mode.manual AND NOT mode.automatic THEN
	_modeToEnum := _E_MainControlMode.manual;
ELSIF mode.automatic AND NOT mode.manual THEN
	_modeToEnum := _E_MainControlMode.automatic;
ELSE
	_modeToEnum := _E_MainControlMode.undefined;
END_IF
END_METHOD

METHOD PROTECTED _plcStateToEnum : _E_MainControlState
VAR_INPUT
	state	: KOSTAL_AF2024_Core_MainControl.I_T_MainControlState;
END_VAR
IF state.PowerOff THEN
	_plcStateToEnum := _E_MainControlState.off;
ELSIF state.RunToHome THEN
	_plcStateToEnum := _E_MainControlState.finish;
ELSIF state.run THEN
	_plcStateToEnum := _E_MainControlState.busy;
ELSIF state.Home THEN
	_plcStateToEnum := _E_MainControlState.ready;
ELSIF state.OnToHome AND NOT state.Home AND NOT state.run AND NOT state.RunToHome THEN
	_plcStateToEnum := _E_MainControlState.calibrate;
ELSIF state.powerOn THEN
	_plcStateToEnum := _E_MainControlState.on;
ELSE
	_plcStateToEnum := _E_MainControlState.off;
END_IF
END_METHOD

METHOD PUBLIC clear
VAR_INPUT
END_VAR


_Name	:= "";

_OnOff.clear();
_runStop.clear();
_RunEmpty.clear();

_Manual.clear();
_Auto.clear();
_Parameters.clear();
_Door.clear();
_Article.clear();

//_statusManual			:= FALSE;
//_statusAuto				:= FALSE;
//_statusData				:= FALSE;
_statusDoor_close	:= FALSE;
_statusDoor_open	:= FALSE;
_statusDoor_safe	:= FALSE;

//_statusOnOff			:= FALSE;
//_statusRun	:= FALSE;
//_statusWorkEmpty	:= FALSE;
//_status.clear();
END_METHOD

METHOD PUBLIC FBmain : BOOL
VAR_INPUT
END_VAR

VAR
END_VAR
IF _mainControl = 0 THEN
	RETURN;
END_IF
IF  _mainControl.Demand = 0 OR _mainControl.Mode = 0 THEN
	RETURN;
END_IF
_buttonHandler();

_mainControlHandler();
END_METHOD

PROPERTY PUBLIC ManualDeviceControl : BOOL
GET
ManualDeviceControl := _manualDeviceControl AND _mainControl.Mode.manual;
END_GET
SET
 _manualDeviceControl := ManualDeviceControl;
END_SET
END_PROPERTY

END_FUNCTION_BLOCK

// MainControl/I_MainControl
(*
Description
===========
| Interface for the main control
*)
INTERFACE I_MainControl

METHOD PUBLIC clear
VAR_INPUT
END_VAR
END_METHOD

END_INTERFACE

// Media/FB_Media
(*

:Author: Martin Hundt <m.hundt@kostal.com>
:Date: 2022-05-05

Function
========
| Adapter for MediaBox on WinHMI 
| File path is set here. Files are stored in WinHMI folder
*)
FUNCTION_BLOCK PUBLIC FB_Media IMPLEMENTS I_Media


VAR

	//****************************************************************************
	//Connector
	//****************************************************************************
	//_connector_FROM_Device	: ST_ARTICLE_FROMDEVICE;	//ST_ARTICLE_FROMDEVICE
	{attribute 'Media_2024_V0'}
	_connector_TO_Device	: _ST_Media_ToDevice;		//ST_ARTICLE_TODEVICE
	//****************************************************************************
	//****************************************************************************
	
	_mediaPath			: T_MEDIA_PATH;
	_standardMediaPath	: T_MEDIA_PATH;
	_showMedia			: BOOL;
END_VAR

//Clear the image or video that was set with SetMedia (display standard image if defined)
METHOD PUBLIC Clear
VAR_INPUT
END_VAR
_mediaPath := '';
END_METHOD

METHOD PUBLIC FBmain : BOOL
IF _mediaPath = '' THEN
	_connector_TO_Device.MediaAddress := _standardMediaPath;
ELSE
	_connector_TO_Device.MediaAddress := _mediaPath;
END_IF

IF _showMedia THEN
	_mediaPath := '';
END_IF

_showMedia := FALSE;
END_METHOD

//Show image or video until it is reset with clear()
//mediaPath is relative to WinHMI location
METHOD PUBLIC SetMedia
VAR_INPUT
	 mediaPath : T_MEDIA_PATH;
END_VAR
_mediaPath := mediaPath;
END_METHOD

//Show image or video as long as this method is called
//mediaPath is relative to WinHMI location
METHOD PUBLIC ShowMedia
VAR_INPUT
	 mediaPath : T_MEDIA_PATH;
END_VAR
_mediaPath := mediaPath;
_showMedia := true;
END_METHOD

//Image or video to show when no other image is defined (optional)
//path is relative to WinHMI location
PROPERTY StandardPath : T_MEDIA_PATH;
GET
StandardPath := _standardMediaPath;
END_GET
SET
_standardMediaPath := StandardPath;
END_SET
END_PROPERTY

END_FUNCTION_BLOCK

// Media/I_Media
(*
Description
===========
| Application interface for MediaBox on WinHMI 
*)
INTERFACE I_Media

//Clear the image or video that was set with SetMedia (display standard image if defined)
METHOD PUBLIC Clear
VAR_INPUT
END_VAR
END_METHOD

//Show image or video until it is reset with clear()
//mediaPath is relative to WinHMI location
METHOD PUBLIC SetMedia
VAR_INPUT
	 mediaPath : T_MEDIA_PATH;
END_VAR
END_METHOD

//Show image or video as long as this method is called
//mediaPath is relative to WinHMI location
METHOD PUBLIC ShowMedia
VAR_INPUT
	 mediaPath : T_MEDIA_PATH;
END_VAR
END_METHOD

//Image or video to show when no other image is defined (optional)
//path is relative to WinHMI location
PROPERTY StandardPath : T_MEDIA_PATH;
GET
END_GET
SET
END_SET
END_PROPERTY

END_INTERFACE

// Parameters/_FB_jsonHandler
FUNCTION_BLOCK _FB_jsonHandler EXTENDS KOSTAL_AF2024_Core_JsonTools._FB_Base_RW

VAR
	_ID			:KOSTAL_AF2024_Core_Settings.T_MaxString_UTF8;
	_Timestamp		:KOSTAL_AF2024_Core_Settings.T_MaxString_UTF8;
	_Values			: ARRAY[1.._NUMBER_OF_VALUES] OF KOSTAL_AF2024_Core_Settings.T_MaxString_UTF8;
END_VAR

VAR CONSTANT
	_ELEMENT_ID			: STRING := 'ID';
	_ELEMENT_TIMESTAMP	: STRING := 'Timestamp';
	_ELEMENT_VALUES		: STRING := 'Values';
	_NUMBER_OF_VALUES 	: USINT := 100;
	
END_VAR

METHOD PUBLIC Clear : BOOL

VAR
	_i: USINT;
END_VAR

_ID			:= '';
_Timestamp 	:= '';

FOR _i := 1 TO _NUMBER_OF_VALUES DO
	_Values[_i]		:= '';
END_FOR


SUPER^.Clear();
END_METHOD

METHOD INTERNAL GetJsonString : T_PARAMETERJSON
VAR
	json : T_PARAMETERJSON;
END_VAR

_parser.CopyDocument(json, SIZEOF(json));

GetJsonString := json;
END_METHOD

METHOD PUBLIC getValue : KOSTAL_AF2024_Core_Settings.T_MaxString_UTF8
VAR_INPUT
	index	: INT;
END_VAR
IF index < 1 OR index > _NUMBER_OF_VALUES THEN
	getValue := 'INVALID';
ELSE
	getValue := _Values[index];
END_IF
END_METHOD

PROPERTY PUBLIC ID :KOSTAL_AF2024_Core_Settings.T_MaxString_UTF8
GET

ID:= _ID;
END_GET
SET

_ID:= ID;
END_SET
END_PROPERTY

PROPERTY PUBLIC NumberOfValues : USINT
GET
NumberOfValues := _NUMBER_OF_VALUES;
END_GET
END_PROPERTY

METHOD PUBLIC setValue : BOOL;
VAR_INPUT
	index	: INT;
	value	: KOSTAL_AF2024_Core_Settings.T_MaxString_UTF8;
END_VAR
IF index < 1 OR index > _NUMBER_OF_VALUES THEN
	setValue :=FALSE;
ELSE
	_Values[index] := value;
	setValue := TRUE;
END_IF
END_METHOD

PROPERTY PUBLIC Timestamp :KOSTAL_AF2024_Core_Settings.T_MaxString_UTF8
GET

Timestamp:= _Timestamp;
END_GET
SET

_Timestamp:= Timestamp;
END_SET
END_PROPERTY

(*
Overwrite to clear your data content before parse content
*)
METHOD PROTECTED _Step_ClearContent
VAR
	_i : USINT;
END_VAR

_ID			:= '';
_Timestamp 	:= '';

FOR _i := 1 TO _NUMBER_OF_VALUES DO
	_Values[_i]		:= '';
END_FOR

SUPER^._Step_ClearContent();
END_METHOD

(*
Overwrite to create your data content
*)
METHOD PROTECTED _Step_CreateContent

VAR
	_jreadArrayElement	: SJsonValue;

	_response 		: KOSTAL_AF2024_Core_Settings.T_MaxString;
	
	//Write
	_jParameterArray		: SJsonValue;
	_i					: UDINT;
END_VAR

_NewDocument();

_parser.AddStringMember(_jDoc, _ELEMENT_ID, _ID);
_parser.AddStringMember(_jDoc, _ELEMENT_TIMESTAMP, _Timestamp);
//_parser.AddArrayMember(_jDoc, _ELEMENT_VALUES, _values);

//Write parameters array
_jParameterArray := _parser.AddArrayMember(_jDoc, _ELEMENT_VALUES,0);
FOR _i:=1 TO _NUMBER_OF_VALUES DO
	_jreadArrayElement := _GetArrayElementByIndex(_jParameterArray, _i, _response);
	_parser.PushbackStringValue(_jParameterArray, _values[_i]);
												
END_FOR


SUPER^._Step_CreateContent();
END_METHOD

(*
Overwrite to parse your data content
*)
METHOD PROTECTED _Step_ParseContent

VAR
	_response: KOSTAL_AF2024_Core_Settings.T_MaxString_UTF8;
	_responseW: KOSTAL_AF2024_Core_Settings.T_MaxString;
	_jValuesArray	: SJsonValue;
	_jArrayElement	: SJsonValue;
	_sParameterValue : STRING;	//Test variable! Remove"
	_i	: USINT;
END_VAR
_ID:= _PARSE_STRING(_jDoc, _ELEMENT_ID, TRUE, _response);

IF _response <> '' THEN ;	END_IF//show error or ...
 

_Timestamp:= _PARSE_STRING(_jDoc, _ELEMENT_TIMESTAMP, TRUE, _response);

IF _response <> '' THEN ;	END_IF//show error or ...


_jValuesArray:= _PARSE_ARRAY(_jDoc, _ELEMENT_VALUES, TRUE, _response);

FOR _i := 1 TO _NUMBER_OF_VALUES DO
	_jArrayElement := _GetArrayElementByIndex(_jValuesArray, (_i-1), _responseW);
	_sParameterValue := _parser.GetString(_jArrayElement);
	_values[_i] := _sParameterValue;
END_FOR



IF _response <> '' THEN ;	END_IF//show error or ...


SUPER^._Step_ParseContent();
END_METHOD

END_FUNCTION_BLOCK

// Parameters/FB_Parameters_Base
(*

:Author: Martin Hundt <m.hundt@kostal.com>
:Date: 2020-12-21

Function
========
Base class to implement WinHMI parameter handlers

Usage
=====
See best practice samples and documentation

*)

FUNCTION_BLOCK FB_Parameters_Base EXTENDS KOSTAL_AF2024_Core_Station.FB_Station_Free IMPLEMENTS  KOSTAL_AF2024_Core_Station.I_Station_Free
VAR
	_mode					: E_DataMode := E_DataMode.ReadFile;
	_init					: BOOL;
	
	//HMI
	_HMI_Station				: FB_Page_Station;
	
	_state					: KOSTAL_AF2024_Core_Process.T_plcState;
	
	
	_jsonHandler			: _FB_jsonHandler;
	_fullQualifiedFile		: KOSTAL_AF2024_Core_Settings.T_MaxString_UTF8;	
	
	//Time
	_I_getTime				: KOSTAL_AF2024_Core_GetSystemTime.I_TimeSource;
	
	//Read File
	_step_readFile			: KOSTAL_AF2024_Core_process.FB_processStep;
	_parameterReadResponse 	: KOSTAL_AF2024_Core_Settings.T_MaxString;
	
	
	//Parameter write parser
	_step_setParameter			: KOSTAL_AF2024_Core_process.FB_processStep;
	
	_setIndex		: USINT;
	_setValue		: T_PARAMETERVALUE;
	_setResponse	: BOOL;
	
	_readFileTimeout		: TON;
	
	//****************************************************************************
	//Connector
	//****************************************************************************
	{attribute 'Parameter_2024_V0'}
	_connector_FROM_Device		: _ST_Parameters_FromDevice;	//ST_DATA_FROMDEVICE
	_connector_TO_Device		: _ST_Parameters_ToDevice;		//ST_DATA_TODEVICE
	//****************************************************************************
END_VAR

VAR CONSTANT
	//NUMBER_OF_PARAMETERS	: INT := 100;
	
	ELEMENT_ID				: STRING := 'ID';
	ELEMENT_TIMESTAMP		: STRING := 'Timestamp';
	ELEMENT_PARAMETERVALUES	: STRING := 'Values';
END_VAR

METHOD PROTECTED _getParameterValue : STRING
VAR_INPUT
	index	: INT;
END_VAR
_getParameterValue := _jsonHandler.getValue(index);
END_METHOD

METHOD _setParameterValue : BOOL;
VAR_INPUT
	Index	: USINT;
	Value	: T_PARAMETERVALUE;
END_VAR
_setIndex := Index;
_setValue := Value;
_mode := E_DataMode.WriteParameter;

_setParameterValue := _setResponse;
END_METHOD

PROPERTY PUBLIC FullQualifiedFile : KOSTAL_AF2024_Core_Settings.T_MaxString_UTF8
GET
FullQualifiedFile := _fullQualifiedFile;
END_GET
SET
_fullQualifiedFile := FullQualifiedFile;
END_SET
END_PROPERTY

METHOD PUBLIC ReloadDataFile
VAR_INPUT
END_VAR
_init := false;
END_METHOD

METHOD INTERNAL _Idle
VAR_INPUT
END_VAR
_step_readFile.init();
_step_setParameter.init();
_setResponse := FALSE;
IF _init THEN
	_message.clear();
	_message.line_01 := "Parameter file loaded successfully";
	_condition.setMessage(KOSTAL_AF2024_Core_process.E_PROCESS_CONDITION_DEFAULT_PRIORITYLEVEL.TEXT_ONLY, _message);
	_state.clear();
	_state.ready := TRUE;
END_IF
END_METHOD

METHOD INTERNAL _readFile : BOOL
VAR

END_VAR
_step_readFile.Header();
_readFile := FALSE;
CASE _step_readFile.actual OF
	0:	//Clear
		_state.clear();
		_state.busy := TRUE;
		_parameterReadResponse := "";
		_readFileTimeout(in:=FALSE);
		_step_readFile.Inc();
		
	
	1:	//Read File
		_readFileTimeout(in:=TRUE, pt:=T#5S);
		IF _jsonHandler.Ex_ReadFile(_fullQualifiedFile) AND _jsonHandler.State.finish AND _jsonHandler.State.pass THEN
			_step_readFile.Inc();
		ELSIF _jsonHandler.State.fail THEN
			_parameterReadResponse := _jsonHandler.State.description;
			_step_readFile.set(10);
		ELSIF _readFileTimeout.Q THEN
			_parameterReadResponse := "Read file timeout";
			_step_readFile.set(10);
		ELSE
			_message.clear();
			_message.line_01 := "Reading parameter file";
			_condition.setMessage(KOSTAL_AF2024_Core_process.E_PROCESS_CONDITION_DEFAULT_PRIORITYLEVEL.MESSAGE, _message);
		END_IF
		
	2:	//Finish
		_readFile := TRUE;
	
	10: //Error
		_message.clear();
		_message.line_01 := "Parameter file invalid";
		_message.line_02 := _parameterReadResponse;
		_condition.setMessage(KOSTAL_AF2024_Core_process.E_PROCESS_CONDITION_DEFAULT_PRIORITYLEVEL.ERROR + 1000, _message);
		_state.clear();
		_state.fail := TRUE;
		_state.description := _parameterReadResponse;
		
		
		
END_CASE
END_METHOD

METHOD PROTECTED _setParaValue : BOOL
VAR
	//read
	_jreadArrayElement	: SJsonValue;

	_response 		: KOSTAL_AF2024_Core_Settings.T_MaxString_UTF8;

	
	//Write
	_jParameterArray		: SJsonValue;
	_i					: UDINT;
	_strJsonParameter	: String(255);
	_exec				: BOOL;
	_sTemp				: STRING;
	
END_VAR
_step_setParameter.Header();
CASE _step_setParameter.actual OF
0:	//Clear
		_state.clear();
		_state.busy := TRUE;
		_parameterReadResponse := "";
		_jsonHandler.setValue(_setIndex, _setValue);
		_readFileTimeout(in:=FALSE);
		_step_setParameter.Inc();
		
	
	1:	//Write File
		_jsonHandler.Timestamp := Tc2_Utilities.SYSTEMTIME_TO_STRING(_I_getTime.GetTimeStruct());
	
		_readFileTimeout(in:=TRUE, pt:=T#5S);
		IF _jsonHandler.Ex_SaveFileAs(_fullQualifiedFile) AND _jsonHandler.State.finish AND _jsonHandler.State.pass THEN
			_step_setParameter.Inc();
		ELSIF _jsonHandler.State.fail THEN
			_parameterReadResponse := _jsonHandler.State.description;
			_step_setParameter.set(10);
		ELSIF _readFileTimeout.Q THEN
			_parameterReadResponse := "Write file timeout";
			_step_setParameter.set(10);
		ELSE
			_message.clear();
			_message.line_01 := "Writing parameter file";
			_condition.setMessage(KOSTAL_AF2024_Core_process.E_PROCESS_CONDITION_DEFAULT_PRIORITYLEVEL.MESSAGE, _message);
		END_IF
		
	2:	//Finish
		_setResponse := TRUE;
		_setParaValue := TRUE;
	
	10: //Error
		_message.clear();
		_message.line_01 := "Parameter file invalid";
		_message.line_02 := _parameterReadResponse;
		_condition.setMessage(KOSTAL_AF2024_Core_process.E_PROCESS_CONDITION_DEFAULT_PRIORITYLEVEL.ERROR + 1000, _message);
		_state.clear();
		_state.fail := TRUE;
		_state.description := _parameterReadResponse;
END_CASE
END_METHOD

METHOD INTERNAL _HMIdefine
VAR
	_i : INT;
END_VAR
//_HMI.linkDataHandler(THIS^);
//_HMI.FBmain();

//=====================================================================================================
// Parameter HMI
//=====================================================================================================
_connector_TO_Device.ParameterValuesJson := _jsonHandler.GetJsonString();

IF _connector_FROM_Device.NewValueTransmit THEN
	IF _setParameterValue(_connector_FROM_Device.SelectedParameter, _connector_FROM_Device.NewValue) THEN
		_connector_TO_Device.NewValueAccept := TRUE;
	END_IF
ELSE
	_connector_TO_Device.NewValueAccept := FALSE;
END_IF


//=====================================================================================================
//Optional station HMI
//=====================================================================================================

_HMI_Station.Name:= "Data Handling";

_HMI_Station.Text.line_01:= _condition.message.line_01;
_HMI_Station.Text.line_02:= _condition.message.line_02;
_HMI_Station.Text.line_03:= _condition.message.line_03;
          
          
_HMI_Station.Button_Escape.Visible	:= _condition.isError();
_HMI_Station.Button_Escape.Text			:= "Reset";
          
_HMI_Station.Status.CopyFrom(_condition);

_HMI_Station.FBmain();
END_METHOD

METHOD PROTECTED _parameterControl : BOOL
VAR_INPUT
END_VAR
//IF _Itext = 0 THEN

//	_message.clear();
//	_message.line_01:= 'Parameter Fail';
//	_message.line_02:= 'Interface _Itext is not linked';

//	_condition.setMessage(4999, _message);
	
IF _I_getTime = 0 THEN

	_message.clear();
	_message.line_01:= "Parameter Fail";
	_message.line_02:= "INTERFACE _I_getTime is NOT linked";

	_condition.setMessage(4999, _message);

ELSE
	
	_parameterControl:= TRUE;

END_IF
END_METHOD

METHOD PROTECTED _resetCondition
VAR_INPUT
END_VAR

IF _condition.isText() THEN
	_condition.clear();
ELSIF _condition.isMessage() THEN
	_condition.clear();
ELSIF _HMI_Station.Button_Escape.Pulse THEN
	_init := false;
	_condition.clear();
END_IF
END_METHOD

METHOD PUBLIC FBmain
VAR
	_i : INT;
END_VAR


//SUPER^.FBmain();

RETURN(NOT _parameterControl());

_HMIdefine();

_jsonHandler.FBmain();

_resetCondition();

IF NOT _init THEN
	_mode := E_DataMode.ReadFile;
END_IF




CASE _mode OF
	E_DataMode.Idle: //Load File
		_Idle();
	E_DataMode.ReadFile:
		IF _readFile()THEN
			_init := TRUE;
		END_IF
	E_DataMode.WriteParameter:
		_setParaValue();
END_CASE

_mode := E_DataMode.Idle;
END_METHOD

METHOD PUBLIC link_I_getTime
VAR_INPUT
	IN : KOSTAL_AF2024_Core_GetSystemTime.I_TimeSource;
END_VAR

_I_getTime:= IN;
END_METHOD

END_FUNCTION_BLOCK

// Project Information/F_GetCompany
// This function has been automatically generated from the project information.
{attribute 'signature_flag' := '1073741824'}
{attribute 'TcGenerated'}
{attribute 'no-analysis'}
FUNCTION F_GetCompany : WSTRING
VAR_INPUT
	
END_VAR

F_GetCompany := "KOSTAL GmbH & Co.KG";

END_FUNCTION

// Project Information/F_GetTitle
// This function has been automatically generated from the project information.
{attribute 'signature_flag' := '1073741824'}
{attribute 'TcGenerated'}
{attribute 'no-analysis'}
FUNCTION F_GetTitle : WSTRING
VAR_INPUT
	
END_VAR

F_GetTitle := "KOSTAL.AF2024.HMI.WinHMI";

END_FUNCTION

// Project Information/F_GetVersion
// This function has been automatically generated from the project information.
{attribute 'signature_flag' := '1073741824'}
{attribute 'TcGenerated'}
{attribute 'no-analysis'}
FUNCTION F_GetVersion : ST_LibVersion
VAR_INPUT
	
END_VAR

F_GetVersion.iMajor := 2;
F_GetVersion.iMinor := 0;
F_GetVersion.iBuild := 0;
F_GetVersion.iRevision := 0;
F_GetVersion.sVersion := '2.0.0.0';
F_GetVersion.nFlags := 0;

END_FUNCTION

// XYZ/FB_page_XYZ
(*

:Author: Martin Hundt <m.hundt@kostal.com>
:Date: 2020-03-09

Function
========
Interface for WinHMI XYZ page

Usage
=====
See best practice samples and documentation

*)


FUNCTION_BLOCK PUBLIC FB_page_XYZ EXTENDS KOSTAL_AF2024_HMI_I_Hmi.FB_page_XYZ


VAR

	//****************************************************************************
	//Connector
	//****************************************************************************
	{attribute 'Page_Xyz_2024_V0'}
	_connector_FROM_Device		: _ST_XYZ_FromDevice;	//ST_3DPAGE_FROMDEVICE
	_connector_TO_Device		: _ST_XYZ_ToDevice;		//ST_3DPAGE_TODEVICE
	//****************************************************************************
	//****************************************************************************

	
	_pulse_forward	: F_TRIG;	
	_pulse_backward	: F_TRIG;	
	_pulse_left		: F_TRIG;	
	_pulse_right	: F_TRIG;	
	_pulse_up		: F_TRIG;	
	_pulse_down		: F_TRIG;	
                             
	_pulse_custom1		: F_TRIG;	
	_pulse_custom2	: F_TRIG;	
	_pulse_custom3		: F_TRIG;	
	_pulse_custom4	: F_TRIG;	
                              
	_pulse_plus		: F_TRIG;	
	_pulse_minus	: F_TRIG;	
	
END_VAR

METHOD PROTECTED _buttonHandler : BOOL
_pulse_forward	(CLK:= _connector_FROM_Device.Button_Forward);
_pulse_backward	(CLK:= _connector_FROM_Device.Button_Backward);
_pulse_left		(CLK:= _connector_FROM_Device.Button_Left);
_pulse_right	(CLK:= _connector_FROM_Device.Button_Right);
_pulse_down		(CLK:= _connector_FROM_Device.Button_Down);
_pulse_up		(CLK:= _connector_FROM_Device.Button_Up);

_pulse_custom1		(CLK:= _connector_FROM_Device.Button_Custom_1);
_pulse_custom2	(CLK:= _connector_FROM_Device.Button_Custom_2);      
_pulse_custom3		(CLK:= _connector_FROM_Device.Button_Custom_3);
_pulse_custom4	(CLK:= _connector_FROM_Device.Button_Custom_4);
      
_pulse_plus		(CLK:= _connector_FROM_Device.Button_StepPlus);
_pulse_minus	(CLK:= _connector_FROM_Device.Button_StepMinus);
END_METHOD

METHOD PROTECTED _fillTextLines
VAR_INPUT
END_VAR

VAR
	_i: INT;
END_VAR
FOR _i:= 1 TO 4 DO
	_connector_TO_Device.Text[_i]:= 	_text[_i];
END_FOR
END_METHOD

METHOD PROTECTED _pageHandler
VAR_INPUT
END_VAR
//Axis (3D)
//TO
_connector_TO_Device.Activate			:= _Activate;
                                                    
_connector_TO_Device.Button_Forward_Active 	:= _Forward.Visible;
_connector_TO_Device.Button_Backward_Active	:= _Backward.Visible;
_connector_TO_Device.Button_Right_Active		:= _Right.Visible;
_connector_TO_Device.Button_Up_Active		:= _Up.Visible;
_connector_TO_Device.Button_Down_Active 		:= _Down.Visible;
_connector_TO_Device.Button_Left_Active		:= _Left.Visible;

_connector_TO_Device.Button_Custom1_Text		:=	_setButton( _Custom.Button_Owner(1));
_connector_TO_Device.Button_Custom2_Text	:= 	_setButton(  _Custom.Button_Owner(2));
_connector_TO_Device.Button_Custom3_Text	:= 	_setButton(  _Custom.Button_Owner(3));
_connector_TO_Device.Button_Custom4_Text		:=	_setButton(  _Custom.Button_Owner(4));

_connector_TO_Device.Button_Plus_Text	:=	_setButton( _Plus);
_connector_TO_Device.Button_Minus_Text	:= 	_setButton( _Minus);

_fillTextLines();

//FROM

_Forward.Sign		:= _connector_FROM_Device.Button_Forward;
_Forward.Pulse	:= _pulse_forward.Q;
_Backward.Sign	:= _connector_FROM_Device.Button_Backward;
_Backward.Pulse	:= _pulse_backward.Q;
 
 
_Left.Sign		:= _connector_FROM_Device.Button_Left;
_Left.Pulse	:= _pulse_left.Q;
 
_Right.Sign	:= _connector_FROM_Device.Button_Right;
_Right.Pulse	:= _pulse_right.Q;
 
_Up.Sign		:= _connector_FROM_Device.Button_Up;
_Up.Pulse	:= _pulse_up.Q;
 
_Down.Sign		:= _connector_FROM_Device.Button_Down;
_Down.Pulse	:= _pulse_down.Q;
 


 _Custom.Button_Owner(1).Sign	:= _connector_FROM_Device.Button_Custom_1;
 _Custom.Button_Owner(1).Pulse	:= _pulse_custom1.Q;

 _Custom.Button_Owner(2).Sign		:= _connector_FROM_Device.Button_Custom_2;
 _Custom.Button_Owner(2).Pulse		:= _pulse_custom2.Q;
 
 _Custom.Button_Owner(3).Sign	:= _connector_FROM_Device.Button_Custom_3;
 _Custom.Button_Owner(3).Pulse	:= _pulse_custom3.Q;
 
 _Custom.Button_Owner(4).Sign	:= _connector_FROM_Device.Button_Custom_4;
 _Custom.Button_Owner(4).Pulse	:= _pulse_custom4.Q;
 
 
_Plus.Sign		:= _connector_FROM_Device.Button_StepPlus;
_Plus.Pulse	:= _pulse_plus.Q;
          
_Minus.Sign	:= _connector_FROM_Device.Button_StepMinus;
_Minus.Pulse	:= _pulse_minus.Q;
END_METHOD

METHOD PROTECTED _setButton : WSTRING

VAR_INPUT
	control	: KOSTAL_AF2024_HMI_Controls.I_T_Button_controlled_Owner;	//KOSTAL_TC3_Controls_button.FB_Button_controlled
END_VAR

IF control.Visible THEN

	IF control.Text = "" THEN
		_setButton:= " ";
	ELSE
		_setButton:= control.Text;
	END_IF

ELSE

	_setButton:= "";

END_IF
END_METHOD

(*
Description
===========
| Method is called automatically
| Do not call manually
*)
METHOD FB_init : BOOL
VAR_INPUT
	bInitRetains : BOOL; // if TRUE, the retain variables are initialized (warm start / cold start)
	bInCopyCode : BOOL;  // if TRUE, the instance afterwards gets moved into the copy code (online change)
END_VAR

VAR
	_index	: INT;	//INT
	x: BOOL;
END_VAR
END_METHOD

METHOD PUBLIC FBmain : BOOL
VAR_INPUT
END_VAR

VAR
END_VAR
_buttonHandler();
_pageHandler();
END_METHOD

END_FUNCTION_BLOCK
